(* IEC 61131-3 sources: s7-to-codesys/tests/POUs/Scenarios/FB_Sequencer_ScenarioTest, 7 files *)

(* ---- FB_Sequencer_ScenarioTest.decl.st ---- *)
// AUTO-GENERATED — не редактировать: s7conv gen-tests, сценарии scenarios/FB_Sequencer.csv
// Правка — в CSV (scenarios/README.md), затем python -m s7conv build-corpus.
// Назначение: тесты поведения сконвертированного FB_Sequencer по сценариям CSV (сценариев: 6, строк: 42):
//             один метод-тест на сценарий, строки — по порядку с моделируемым временем GVL_S7Clock.
//             Ожидаемые значения — из CSV (эталонные модели по описанию логики блока), не из
//             результата конвертации.
// Автор:      s7conv 0.1.0 (сгенерировано)
// Версия:     не указана
// Документ:   scenarios/README.md, docs/methodology.md, раздел «Проверка поведения»
FUNCTION_BLOCK FB_Sequencer_ScenarioTest EXTENDS coUnit.FB_TestSuite
VAR
    fbFullCycle : FB_Sequencer;  // свой экземпляр на сценарий
    xFullCycleDone : BOOL;  // сценарий выполнен (выполняется один раз)
    fbDrainTimeout : FB_Sequencer;  // свой экземпляр на сценарий
    xDrainTimeoutDone : BOOL;  // сценарий выполнен (выполняется один раз)
    fbAbortByStop : FB_Sequencer;  // свой экземпляр на сценарий
    xAbortByStopDone : BOOL;  // сценарий выполнен (выполняется один раз)
    fbPermissiveMissing : FB_Sequencer;  // свой экземпляр на сценарий
    xPermissiveMissingDone : BOOL;  // сценарий выполнен (выполняется один раз)
    fbDrainTimeoutBoundary : FB_Sequencer;  // свой экземпляр на сценарий
    xDrainTimeoutBoundaryDone : BOOL;  // сценарий выполнен (выполняется один раз)
    fbRefillTimeoutBoundary : FB_Sequencer;  // свой экземпляр на сценарий
    xRefillTimeoutBoundaryDone : BOOL;  // сценарий выполнен (выполняется один раз)
END_VAR

(* ---- AbortByStop.method.impl.st ---- *)
// AUTO-GENERATED — не редактировать: scenarios/FB_Sequencer.csv, сценарий AbortByStop
coUnit.TEST('AbortByStop');
IF NOT xAbortByStopDone THEN
    xAbortByStopDone := TRUE;
    GVL_S7Clock.xSimulation := TRUE;

    // #1, t = 0 мс — ожидание
    GVL_S7Clock.tSimNow := T#0MS;
    fbAbortByStop.start := FALSE;
    fbAbortByStop.stop := FALSE;
    fbAbortByStop.permissive := TRUE;
    fbAbortByStop.levelLow := FALSE;
    fbAbortByStop.levelHigh := FALSE;
    fbAbortByStop.reset := FALSE;
    fbAbortByStop.drainTimeout := T#60000MS;
    fbAbortByStop.airTime := T#30000MS;
    fbAbortByStop.washTime := T#40000MS;
    fbAbortByStop.refillTimeout := T#90000MS;
    fbAbortByStop();
    AssertEquals_INT(Expected := 0, Actual := fbAbortByStop.stepNo, Message := 'AbortByStop#1 stepNo');
    AssertEquals_BOOL(Expected := FALSE, Actual := fbAbortByStop.drainValve, Message := 'AbortByStop#1 drainValve');
    AssertEquals_BOOL(Expected := FALSE, Actual := fbAbortByStop.airBlower, Message := 'AbortByStop#1 airBlower');
    AssertEquals_BOOL(Expected := FALSE, Actual := fbAbortByStop.washPump, Message := 'AbortByStop#1 washPump');
    AssertEquals_BOOL(Expected := FALSE, Actual := fbAbortByStop.inletValve, Message := 'AbortByStop#1 inletValve');
    AssertEquals_BOOL(Expected := FALSE, Actual := fbAbortByStop.busy, Message := 'AbortByStop#1 busy');
    AssertEquals_BOOL(Expected := FALSE, Actual := fbAbortByStop.fault, Message := 'AbortByStop#1 fault');
    AssertEquals_INT(Expected := 0, Actual := fbAbortByStop.faultStep, Message := 'AbortByStop#1 faultStep');
    AssertEquals_DINT(Expected := 0, Actual := fbAbortByStop.cycleCount, Message := 'AbortByStop#1 cycleCount');
    AssertEquals_STRING(Expected := 'IDLE', Actual := fbAbortByStop.stepText, Message := 'AbortByStop#1 stepText');

    // #2, t = 1000 мс — пуск: опорожнение
    GVL_S7Clock.tSimNow := T#1000MS;
    fbAbortByStop.start := TRUE;
    fbAbortByStop();
    AssertEquals_INT(Expected := 10, Actual := fbAbortByStop.stepNo, Message := 'AbortByStop#2 stepNo');
    AssertEquals_BOOL(Expected := TRUE, Actual := fbAbortByStop.drainValve, Message := 'AbortByStop#2 drainValve');
    AssertEquals_BOOL(Expected := FALSE, Actual := fbAbortByStop.airBlower, Message := 'AbortByStop#2 airBlower');
    AssertEquals_BOOL(Expected := FALSE, Actual := fbAbortByStop.washPump, Message := 'AbortByStop#2 washPump');
    AssertEquals_BOOL(Expected := FALSE, Actual := fbAbortByStop.inletValve, Message := 'AbortByStop#2 inletValve');
    AssertEquals_BOOL(Expected := TRUE, Actual := fbAbortByStop.busy, Message := 'AbortByStop#2 busy');
    AssertEquals_BOOL(Expected := FALSE, Actual := fbAbortByStop.fault, Message := 'AbortByStop#2 fault');
    AssertEquals_INT(Expected := 0, Actual := fbAbortByStop.faultStep, Message := 'AbortByStop#2 faultStep');
    AssertEquals_DINT(Expected := 0, Actual := fbAbortByStop.cycleCount, Message := 'AbortByStop#2 cycleCount');
    AssertEquals_STRING(Expected := 'DRAIN', Actual := fbAbortByStop.stepText, Message := 'AbortByStop#2 stepText');

    // #3, t = 5000 мс — продувка с 5.0 с
    GVL_S7Clock.tSimNow := T#5000MS;
    fbAbortByStop.start := FALSE;
    fbAbortByStop.levelLow := TRUE;
    fbAbortByStop();
    AssertEquals_INT(Expected := 20, Actual := fbAbortByStop.stepNo, Message := 'AbortByStop#3 stepNo');
    AssertEquals_BOOL(Expected := FALSE, Actual := fbAbortByStop.drainValve, Message := 'AbortByStop#3 drainValve');
    AssertEquals_BOOL(Expected := TRUE, Actual := fbAbortByStop.airBlower, Message := 'AbortByStop#3 airBlower');
    AssertEquals_BOOL(Expected := FALSE, Actual := fbAbortByStop.washPump, Message := 'AbortByStop#3 washPump');
    AssertEquals_BOOL(Expected := FALSE, Actual := fbAbortByStop.inletValve, Message := 'AbortByStop#3 inletValve');
    AssertEquals_BOOL(Expected := TRUE, Actual := fbAbortByStop.busy, Message := 'AbortByStop#3 busy');
    AssertEquals_BOOL(Expected := FALSE, Actual := fbAbortByStop.fault, Message := 'AbortByStop#3 fault');
    AssertEquals_INT(Expected := 0, Actual := fbAbortByStop.faultStep, Message := 'AbortByStop#3 faultStep');
    AssertEquals_DINT(Expected := 0, Actual := fbAbortByStop.cycleCount, Message := 'AbortByStop#3 cycleCount');
    AssertEquals_STRING(Expected := 'AIR SCOUR', Actual := fbAbortByStop.stepText, Message := 'AbortByStop#3 stepText');

    // #4, t = 10000 мс — прерывание: ожидание, без аварии и без счёта
    GVL_S7Clock.tSimNow := T#10000MS;
    fbAbortByStop.stop := TRUE;
    fbAbortByStop();
    AssertEquals_INT(Expected := 0, Actual := fbAbortByStop.stepNo, Message := 'AbortByStop#4 stepNo');
    AssertEquals_BOOL(Expected := FALSE, Actual := fbAbortByStop.drainValve, Message := 'AbortByStop#4 drainValve');
    AssertEquals_BOOL(Expected := FALSE, Actual := fbAbortByStop.airBlower, Message := 'AbortByStop#4 airBlower');
    AssertEquals_BOOL(Expected := FALSE, Actual := fbAbortByStop.washPump, Message := 'AbortByStop#4 washPump');
    AssertEquals_BOOL(Expected := FALSE, Actual := fbAbortByStop.inletValve, Message := 'AbortByStop#4 inletValve');
    AssertEquals_BOOL(Expected := FALSE, Actual := fbAbortByStop.busy, Message := 'AbortByStop#4 busy');
    AssertEquals_BOOL(Expected := FALSE, Actual := fbAbortByStop.fault, Message := 'AbortByStop#4 fault');
    AssertEquals_INT(Expected := 0, Actual := fbAbortByStop.faultStep, Message := 'AbortByStop#4 faultStep');
    AssertEquals_DINT(Expected := 0, Actual := fbAbortByStop.cycleCount, Message := 'AbortByStop#4 cycleCount');
    AssertEquals_STRING(Expected := 'IDLE', Actual := fbAbortByStop.stepText, Message := 'AbortByStop#4 stepText');

    // #5, t = 11000 мс — фронт start при stop: не запускается
    GVL_S7Clock.tSimNow := T#11000MS;
    fbAbortByStop.start := TRUE;
    fbAbortByStop();
    AssertEquals_INT(Expected := 0, Actual := fbAbortByStop.stepNo, Message := 'AbortByStop#5 stepNo');
    AssertEquals_BOOL(Expected := FALSE, Actual := fbAbortByStop.drainValve, Message := 'AbortByStop#5 drainValve');
    AssertEquals_BOOL(Expected := FALSE, Actual := fbAbortByStop.airBlower, Message := 'AbortByStop#5 airBlower');
    AssertEquals_BOOL(Expected := FALSE, Actual := fbAbortByStop.washPump, Message := 'AbortByStop#5 washPump');
    AssertEquals_BOOL(Expected := FALSE, Actual := fbAbortByStop.inletValve, Message := 'AbortByStop#5 inletValve');
    AssertEquals_BOOL(Expected := FALSE, Actual := fbAbortByStop.busy, Message := 'AbortByStop#5 busy');
    AssertEquals_BOOL(Expected := FALSE, Actual := fbAbortByStop.fault, Message := 'AbortByStop#5 fault');
    AssertEquals_INT(Expected := 0, Actual := fbAbortByStop.faultStep, Message := 'AbortByStop#5 faultStep');
    AssertEquals_DINT(Expected := 0, Actual := fbAbortByStop.cycleCount, Message := 'AbortByStop#5 cycleCount');
    AssertEquals_STRING(Expected := 'IDLE', Actual := fbAbortByStop.stepText, Message := 'AbortByStop#5 stepText');

    // #6, t = 12000 мс — stop снят
    GVL_S7Clock.tSimNow := T#12000MS;
    fbAbortByStop.start := FALSE;
    fbAbortByStop.stop := FALSE;
    fbAbortByStop();
    AssertEquals_INT(Expected := 0, Actual := fbAbortByStop.stepNo, Message := 'AbortByStop#6 stepNo');
    AssertEquals_BOOL(Expected := FALSE, Actual := fbAbortByStop.drainValve, Message := 'AbortByStop#6 drainValve');
    AssertEquals_BOOL(Expected := FALSE, Actual := fbAbortByStop.airBlower, Message := 'AbortByStop#6 airBlower');
    AssertEquals_BOOL(Expected := FALSE, Actual := fbAbortByStop.washPump, Message := 'AbortByStop#6 washPump');
    AssertEquals_BOOL(Expected := FALSE, Actual := fbAbortByStop.inletValve, Message := 'AbortByStop#6 inletValve');
    AssertEquals_BOOL(Expected := FALSE, Actual := fbAbortByStop.busy, Message := 'AbortByStop#6 busy');
    AssertEquals_BOOL(Expected := FALSE, Actual := fbAbortByStop.fault, Message := 'AbortByStop#6 fault');
    AssertEquals_INT(Expected := 0, Actual := fbAbortByStop.faultStep, Message := 'AbortByStop#6 faultStep');
    AssertEquals_DINT(Expected := 0, Actual := fbAbortByStop.cycleCount, Message := 'AbortByStop#6 cycleCount');
    AssertEquals_STRING(Expected := 'IDLE', Actual := fbAbortByStop.stepText, Message := 'AbortByStop#6 stepText');

    // #7, t = 13000 мс — новый фронт start: опорожнение
    GVL_S7Clock.tSimNow := T#13000MS;
    fbAbortByStop.start := TRUE;
    fbAbortByStop();
    AssertEquals_INT(Expected := 10, Actual := fbAbortByStop.stepNo, Message := 'AbortByStop#7 stepNo');
    AssertEquals_BOOL(Expected := TRUE, Actual := fbAbortByStop.drainValve, Message := 'AbortByStop#7 drainValve');
    AssertEquals_BOOL(Expected := FALSE, Actual := fbAbortByStop.airBlower, Message := 'AbortByStop#7 airBlower');
    AssertEquals_BOOL(Expected := FALSE, Actual := fbAbortByStop.washPump, Message := 'AbortByStop#7 washPump');
    AssertEquals_BOOL(Expected := FALSE, Actual := fbAbortByStop.inletValve, Message := 'AbortByStop#7 inletValve');
    AssertEquals_BOOL(Expected := TRUE, Actual := fbAbortByStop.busy, Message := 'AbortByStop#7 busy');
    AssertEquals_BOOL(Expected := FALSE, Actual := fbAbortByStop.fault, Message := 'AbortByStop#7 fault');
    AssertEquals_INT(Expected := 0, Actual := fbAbortByStop.faultStep, Message := 'AbortByStop#7 faultStep');
    AssertEquals_DINT(Expected := 0, Actual := fbAbortByStop.cycleCount, Message := 'AbortByStop#7 cycleCount');
    AssertEquals_STRING(Expected := 'DRAIN', Actual := fbAbortByStop.stepText, Message := 'AbortByStop#7 stepText');

    GVL_S7Clock.xSimulation := FALSE;
END_IF
coUnit.TEST_FINISHED();

(* ---- DrainTimeout.method.impl.st ---- *)
// AUTO-GENERATED — не редактировать: scenarios/FB_Sequencer.csv, сценарий DrainTimeout
coUnit.TEST('DrainTimeout');
IF NOT xDrainTimeoutDone THEN
    xDrainTimeoutDone := TRUE;
    GVL_S7Clock.xSimulation := TRUE;

    // #1, t = 0 мс — ожидание
    GVL_S7Clock.tSimNow := T#0MS;
    fbDrainTimeout.start := FALSE;
    fbDrainTimeout.stop := FALSE;
    fbDrainTimeout.permissive := TRUE;
    fbDrainTimeout.levelLow := FALSE;
    fbDrainTimeout.levelHigh := FALSE;
    fbDrainTimeout.reset := FALSE;
    fbDrainTimeout.drainTimeout := T#60000MS;
    fbDrainTimeout.airTime := T#30000MS;
    fbDrainTimeout.washTime := T#40000MS;
    fbDrainTimeout.refillTimeout := T#90000MS;
    fbDrainTimeout();
    AssertEquals_INT(Expected := 0, Actual := fbDrainTimeout.stepNo, Message := 'DrainTimeout#1 stepNo');
    AssertEquals_BOOL(Expected := FALSE, Actual := fbDrainTimeout.drainValve, Message := 'DrainTimeout#1 drainValve');
    AssertEquals_BOOL(Expected := FALSE, Actual := fbDrainTimeout.airBlower, Message := 'DrainTimeout#1 airBlower');
    AssertEquals_BOOL(Expected := FALSE, Actual := fbDrainTimeout.washPump, Message := 'DrainTimeout#1 washPump');
    AssertEquals_BOOL(Expected := FALSE, Actual := fbDrainTimeout.inletValve, Message := 'DrainTimeout#1 inletValve');
    AssertEquals_BOOL(Expected := FALSE, Actual := fbDrainTimeout.busy, Message := 'DrainTimeout#1 busy');
    AssertEquals_BOOL(Expected := FALSE, Actual := fbDrainTimeout.fault, Message := 'DrainTimeout#1 fault');
    AssertEquals_INT(Expected := 0, Actual := fbDrainTimeout.faultStep, Message := 'DrainTimeout#1 faultStep');
    AssertEquals_DINT(Expected := 0, Actual := fbDrainTimeout.cycleCount, Message := 'DrainTimeout#1 cycleCount');
    AssertEquals_STRING(Expected := 'IDLE', Actual := fbDrainTimeout.stepText, Message := 'DrainTimeout#1 stepText');

    // #2, t = 1000 мс — пуск: опорожнение с 1.0 с
    GVL_S7Clock.tSimNow := T#1000MS;
    fbDrainTimeout.start := TRUE;
    fbDrainTimeout();
    AssertEquals_INT(Expected := 10, Actual := fbDrainTimeout.stepNo, Message := 'DrainTimeout#2 stepNo');
    AssertEquals_BOOL(Expected := TRUE, Actual := fbDrainTimeout.drainValve, Message := 'DrainTimeout#2 drainValve');
    AssertEquals_BOOL(Expected := FALSE, Actual := fbDrainTimeout.airBlower, Message := 'DrainTimeout#2 airBlower');
    AssertEquals_BOOL(Expected := FALSE, Actual := fbDrainTimeout.washPump, Message := 'DrainTimeout#2 washPump');
    AssertEquals_BOOL(Expected := FALSE, Actual := fbDrainTimeout.inletValve, Message := 'DrainTimeout#2 inletValve');
    AssertEquals_BOOL(Expected := TRUE, Actual := fbDrainTimeout.busy, Message := 'DrainTimeout#2 busy');
    AssertEquals_BOOL(Expected := FALSE, Actual := fbDrainTimeout.fault, Message := 'DrainTimeout#2 fault');
    AssertEquals_INT(Expected := 0, Actual := fbDrainTimeout.faultStep, Message := 'DrainTimeout#2 faultStep');
    AssertEquals_DINT(Expected := 0, Actual := fbDrainTimeout.cycleCount, Message := 'DrainTimeout#2 cycleCount');
    AssertEquals_STRING(Expected := 'DRAIN', Actual := fbDrainTimeout.stepText, Message := 'DrainTimeout#2 stepText');

    // #3, t = 60800 мс — 59.8 с < 60 с: опорожнение
    GVL_S7Clock.tSimNow := T#60800MS;
    fbDrainTimeout.start := FALSE;
    fbDrainTimeout();
    AssertEquals_INT(Expected := 10, Actual := fbDrainTimeout.stepNo, Message := 'DrainTimeout#3 stepNo');
    AssertEquals_BOOL(Expected := TRUE, Actual := fbDrainTimeout.drainValve, Message := 'DrainTimeout#3 drainValve');
    AssertEquals_BOOL(Expected := FALSE, Actual := fbDrainTimeout.airBlower, Message := 'DrainTimeout#3 airBlower');
    AssertEquals_BOOL(Expected := FALSE, Actual := fbDrainTimeout.washPump, Message := 'DrainTimeout#3 washPump');
    AssertEquals_BOOL(Expected := FALSE, Actual := fbDrainTimeout.inletValve, Message := 'DrainTimeout#3 inletValve');
    AssertEquals_BOOL(Expected := TRUE, Actual := fbDrainTimeout.busy, Message := 'DrainTimeout#3 busy');
    AssertEquals_BOOL(Expected := FALSE, Actual := fbDrainTimeout.fault, Message := 'DrainTimeout#3 fault');
    AssertEquals_INT(Expected := 0, Actual := fbDrainTimeout.faultStep, Message := 'DrainTimeout#3 faultStep');
    AssertEquals_DINT(Expected := 0, Actual := fbDrainTimeout.cycleCount, Message := 'DrainTimeout#3 cycleCount');
    AssertEquals_STRING(Expected := 'DRAIN', Actual := fbDrainTimeout.stepText, Message := 'DrainTimeout#3 stepText');

    // #4, t = 61200 мс — 60.2 с: авария на шаге 10, всё закрыто
    GVL_S7Clock.tSimNow := T#61200MS;
    fbDrainTimeout();
    AssertEquals_INT(Expected := 90, Actual := fbDrainTimeout.stepNo, Message := 'DrainTimeout#4 stepNo');
    AssertEquals_BOOL(Expected := FALSE, Actual := fbDrainTimeout.drainValve, Message := 'DrainTimeout#4 drainValve');
    AssertEquals_BOOL(Expected := FALSE, Actual := fbDrainTimeout.airBlower, Message := 'DrainTimeout#4 airBlower');
    AssertEquals_BOOL(Expected := FALSE, Actual := fbDrainTimeout.washPump, Message := 'DrainTimeout#4 washPump');
    AssertEquals_BOOL(Expected := FALSE, Actual := fbDrainTimeout.inletValve, Message := 'DrainTimeout#4 inletValve');
    AssertEquals_BOOL(Expected := FALSE, Actual := fbDrainTimeout.busy, Message := 'DrainTimeout#4 busy');
    AssertEquals_BOOL(Expected := TRUE, Actual := fbDrainTimeout.fault, Message := 'DrainTimeout#4 fault');
    AssertEquals_INT(Expected := 10, Actual := fbDrainTimeout.faultStep, Message := 'DrainTimeout#4 faultStep');
    AssertEquals_DINT(Expected := 0, Actual := fbDrainTimeout.cycleCount, Message := 'DrainTimeout#4 cycleCount');
    AssertEquals_STRING(Expected := 'FAULT', Actual := fbDrainTimeout.stepText, Message := 'DrainTimeout#4 stepText');

    // #5, t = 65000 мс — пуск во время аварии не действует
    GVL_S7Clock.tSimNow := T#65000MS;
    fbDrainTimeout.start := TRUE;
    fbDrainTimeout();
    AssertEquals_INT(Expected := 90, Actual := fbDrainTimeout.stepNo, Message := 'DrainTimeout#5 stepNo');
    AssertEquals_BOOL(Expected := FALSE, Actual := fbDrainTimeout.drainValve, Message := 'DrainTimeout#5 drainValve');
    AssertEquals_BOOL(Expected := FALSE, Actual := fbDrainTimeout.airBlower, Message := 'DrainTimeout#5 airBlower');
    AssertEquals_BOOL(Expected := FALSE, Actual := fbDrainTimeout.washPump, Message := 'DrainTimeout#5 washPump');
    AssertEquals_BOOL(Expected := FALSE, Actual := fbDrainTimeout.inletValve, Message := 'DrainTimeout#5 inletValve');
    AssertEquals_BOOL(Expected := FALSE, Actual := fbDrainTimeout.busy, Message := 'DrainTimeout#5 busy');
    AssertEquals_BOOL(Expected := TRUE, Actual := fbDrainTimeout.fault, Message := 'DrainTimeout#5 fault');
    AssertEquals_INT(Expected := 10, Actual := fbDrainTimeout.faultStep, Message := 'DrainTimeout#5 faultStep');
    AssertEquals_DINT(Expected := 0, Actual := fbDrainTimeout.cycleCount, Message := 'DrainTimeout#5 cycleCount');
    AssertEquals_STRING(Expected := 'FAULT', Actual := fbDrainTimeout.stepText, Message := 'DrainTimeout#5 stepText');

    // #6, t = 70000 мс — сброс: ожидание, faultStep 0
    GVL_S7Clock.tSimNow := T#70000MS;
    fbDrainTimeout.start := FALSE;
    fbDrainTimeout.reset := TRUE;
    fbDrainTimeout();
    AssertEquals_INT(Expected := 0, Actual := fbDrainTimeout.stepNo, Message := 'DrainTimeout#6 stepNo');
    AssertEquals_BOOL(Expected := FALSE, Actual := fbDrainTimeout.drainValve, Message := 'DrainTimeout#6 drainValve');
    AssertEquals_BOOL(Expected := FALSE, Actual := fbDrainTimeout.airBlower, Message := 'DrainTimeout#6 airBlower');
    AssertEquals_BOOL(Expected := FALSE, Actual := fbDrainTimeout.washPump, Message := 'DrainTimeout#6 washPump');
    AssertEquals_BOOL(Expected := FALSE, Actual := fbDrainTimeout.inletValve, Message := 'DrainTimeout#6 inletValve');
    AssertEquals_BOOL(Expected := FALSE, Actual := fbDrainTimeout.busy, Message := 'DrainTimeout#6 busy');
    AssertEquals_BOOL(Expected := FALSE, Actual := fbDrainTimeout.fault, Message := 'DrainTimeout#6 fault');
    AssertEquals_INT(Expected := 0, Actual := fbDrainTimeout.faultStep, Message := 'DrainTimeout#6 faultStep');
    AssertEquals_DINT(Expected := 0, Actual := fbDrainTimeout.cycleCount, Message := 'DrainTimeout#6 cycleCount');
    AssertEquals_STRING(Expected := 'IDLE', Actual := fbDrainTimeout.stepText, Message := 'DrainTimeout#6 stepText');

    // #7, t = 71000 мс — ожидание
    GVL_S7Clock.tSimNow := T#71000MS;
    fbDrainTimeout.reset := FALSE;
    fbDrainTimeout();
    AssertEquals_INT(Expected := 0, Actual := fbDrainTimeout.stepNo, Message := 'DrainTimeout#7 stepNo');
    AssertEquals_BOOL(Expected := FALSE, Actual := fbDrainTimeout.drainValve, Message := 'DrainTimeout#7 drainValve');
    AssertEquals_BOOL(Expected := FALSE, Actual := fbDrainTimeout.airBlower, Message := 'DrainTimeout#7 airBlower');
    AssertEquals_BOOL(Expected := FALSE, Actual := fbDrainTimeout.washPump, Message := 'DrainTimeout#7 washPump');
    AssertEquals_BOOL(Expected := FALSE, Actual := fbDrainTimeout.inletValve, Message := 'DrainTimeout#7 inletValve');
    AssertEquals_BOOL(Expected := FALSE, Actual := fbDrainTimeout.busy, Message := 'DrainTimeout#7 busy');
    AssertEquals_BOOL(Expected := FALSE, Actual := fbDrainTimeout.fault, Message := 'DrainTimeout#7 fault');
    AssertEquals_INT(Expected := 0, Actual := fbDrainTimeout.faultStep, Message := 'DrainTimeout#7 faultStep');
    AssertEquals_DINT(Expected := 0, Actual := fbDrainTimeout.cycleCount, Message := 'DrainTimeout#7 cycleCount');
    AssertEquals_STRING(Expected := 'IDLE', Actual := fbDrainTimeout.stepText, Message := 'DrainTimeout#7 stepText');

    GVL_S7Clock.xSimulation := FALSE;
END_IF
coUnit.TEST_FINISHED();

(* ---- DrainTimeoutBoundary.method.impl.st ---- *)
// AUTO-GENERATED — не редактировать: scenarios/FB_Sequencer.csv, сценарий DrainTimeoutBoundary
coUnit.TEST('DrainTimeoutBoundary');
IF NOT xDrainTimeoutBoundaryDone THEN
    xDrainTimeoutBoundaryDone := TRUE;
    GVL_S7Clock.xSimulation := TRUE;

    // #1, t = 0 мс — пуск в первом вызове: опорожнение с 0 с
    GVL_S7Clock.tSimNow := T#0MS;
    fbDrainTimeoutBoundary.start := TRUE;
    fbDrainTimeoutBoundary.stop := FALSE;
    fbDrainTimeoutBoundary.permissive := TRUE;
    fbDrainTimeoutBoundary.levelLow := FALSE;
    fbDrainTimeoutBoundary.levelHigh := FALSE;
    fbDrainTimeoutBoundary.reset := FALSE;
    fbDrainTimeoutBoundary.drainTimeout := T#60000MS;
    fbDrainTimeoutBoundary.airTime := T#30000MS;
    fbDrainTimeoutBoundary.washTime := T#40000MS;
    fbDrainTimeoutBoundary.refillTimeout := T#90000MS;
    fbDrainTimeoutBoundary();
    AssertEquals_INT(Expected := 10,
                     Actual := fbDrainTimeoutBoundary.stepNo,
                     Message := 'DrainTimeoutBoundary#1 stepNo');
    AssertEquals_BOOL(Expected := TRUE,
                      Actual := fbDrainTimeoutBoundary.drainValve,
                      Message := 'DrainTimeoutBoundary#1 drainValve');
    AssertEquals_BOOL(Expected := FALSE,
                      Actual := fbDrainTimeoutBoundary.airBlower,
                      Message := 'DrainTimeoutBoundary#1 airBlower');
    AssertEquals_BOOL(Expected := FALSE,
                      Actual := fbDrainTimeoutBoundary.washPump,
                      Message := 'DrainTimeoutBoundary#1 washPump');
    AssertEquals_BOOL(Expected := FALSE,
                      Actual := fbDrainTimeoutBoundary.inletValve,
                      Message := 'DrainTimeoutBoundary#1 inletValve');
    AssertEquals_BOOL(Expected := TRUE,
                      Actual := fbDrainTimeoutBoundary.busy,
                      Message := 'DrainTimeoutBoundary#1 busy');
    AssertEquals_BOOL(Expected := FALSE,
                      Actual := fbDrainTimeoutBoundary.fault,
                      Message := 'DrainTimeoutBoundary#1 fault');
    AssertEquals_INT(Expected := 0,
                     Actual := fbDrainTimeoutBoundary.faultStep,
                     Message := 'DrainTimeoutBoundary#1 faultStep');
    AssertEquals_DINT(Expected := 0,
                      Actual := fbDrainTimeoutBoundary.cycleCount,
                      Message := 'DrainTimeoutBoundary#1 cycleCount');
    AssertEquals_STRING(Expected := 'DRAIN',
                        Actual := fbDrainTimeoutBoundary.stepText,
                        Message := 'DrainTimeoutBoundary#1 stepText');

    // #2, t = 59800 мс — 59.8 с: опорожнение
    GVL_S7Clock.tSimNow := T#59800MS;
    fbDrainTimeoutBoundary.start := FALSE;
    fbDrainTimeoutBoundary();
    AssertEquals_INT(Expected := 10,
                     Actual := fbDrainTimeoutBoundary.stepNo,
                     Message := 'DrainTimeoutBoundary#2 stepNo');
    AssertEquals_BOOL(Expected := TRUE,
                      Actual := fbDrainTimeoutBoundary.drainValve,
                      Message := 'DrainTimeoutBoundary#2 drainValve');
    AssertEquals_BOOL(Expected := FALSE,
                      Actual := fbDrainTimeoutBoundary.airBlower,
                      Message := 'DrainTimeoutBoundary#2 airBlower');
    AssertEquals_BOOL(Expected := FALSE,
                      Actual := fbDrainTimeoutBoundary.washPump,
                      Message := 'DrainTimeoutBoundary#2 washPump');
    AssertEquals_BOOL(Expected := FALSE,
                      Actual := fbDrainTimeoutBoundary.inletValve,
                      Message := 'DrainTimeoutBoundary#2 inletValve');
    AssertEquals_BOOL(Expected := TRUE,
                      Actual := fbDrainTimeoutBoundary.busy,
                      Message := 'DrainTimeoutBoundary#2 busy');
    AssertEquals_BOOL(Expected := FALSE,
                      Actual := fbDrainTimeoutBoundary.fault,
                      Message := 'DrainTimeoutBoundary#2 fault');
    AssertEquals_INT(Expected := 0,
                     Actual := fbDrainTimeoutBoundary.faultStep,
                     Message := 'DrainTimeoutBoundary#2 faultStep');
    AssertEquals_DINT(Expected := 0,
                      Actual := fbDrainTimeoutBoundary.cycleCount,
                      Message := 'DrainTimeoutBoundary#2 cycleCount');
    AssertEquals_STRING(Expected := 'DRAIN',
                        Actual := fbDrainTimeoutBoundary.stepText,
                        Message := 'DrainTimeoutBoundary#2 stepText');

    // #3, t = 60000 мс, на пороге таймера — 60.0 с = drainTimeout: авария
    GVL_S7Clock.tSimNow := T#60000MS;
    fbDrainTimeoutBoundary();
    AssertEquals_INT(Expected := 90,
                     Actual := fbDrainTimeoutBoundary.stepNo,
                     Message := 'DrainTimeoutBoundary#3 stepNo');
    AssertEquals_BOOL(Expected := FALSE,
                      Actual := fbDrainTimeoutBoundary.drainValve,
                      Message := 'DrainTimeoutBoundary#3 drainValve');
    AssertEquals_BOOL(Expected := FALSE,
                      Actual := fbDrainTimeoutBoundary.airBlower,
                      Message := 'DrainTimeoutBoundary#3 airBlower');
    AssertEquals_BOOL(Expected := FALSE,
                      Actual := fbDrainTimeoutBoundary.washPump,
                      Message := 'DrainTimeoutBoundary#3 washPump');
    AssertEquals_BOOL(Expected := FALSE,
                      Actual := fbDrainTimeoutBoundary.inletValve,
                      Message := 'DrainTimeoutBoundary#3 inletValve');
    AssertEquals_BOOL(Expected := FALSE,
                      Actual := fbDrainTimeoutBoundary.busy,
                      Message := 'DrainTimeoutBoundary#3 busy');
    AssertEquals_BOOL(Expected := TRUE,
                      Actual := fbDrainTimeoutBoundary.fault,
                      Message := 'DrainTimeoutBoundary#3 fault');
    AssertEquals_INT(Expected := 10,
                     Actual := fbDrainTimeoutBoundary.faultStep,
                     Message := 'DrainTimeoutBoundary#3 faultStep');
    AssertEquals_DINT(Expected := 0,
                      Actual := fbDrainTimeoutBoundary.cycleCount,
                      Message := 'DrainTimeoutBoundary#3 cycleCount');
    AssertEquals_STRING(Expected := 'FAULT',
                        Actual := fbDrainTimeoutBoundary.stepText,
                        Message := 'DrainTimeoutBoundary#3 stepText');

    // #4, t = 60200 мс — авария
    GVL_S7Clock.tSimNow := T#60200MS;
    fbDrainTimeoutBoundary();
    AssertEquals_INT(Expected := 90,
                     Actual := fbDrainTimeoutBoundary.stepNo,
                     Message := 'DrainTimeoutBoundary#4 stepNo');
    AssertEquals_BOOL(Expected := FALSE,
                      Actual := fbDrainTimeoutBoundary.drainValve,
                      Message := 'DrainTimeoutBoundary#4 drainValve');
    AssertEquals_BOOL(Expected := FALSE,
                      Actual := fbDrainTimeoutBoundary.airBlower,
                      Message := 'DrainTimeoutBoundary#4 airBlower');
    AssertEquals_BOOL(Expected := FALSE,
                      Actual := fbDrainTimeoutBoundary.washPump,
                      Message := 'DrainTimeoutBoundary#4 washPump');
    AssertEquals_BOOL(Expected := FALSE,
                      Actual := fbDrainTimeoutBoundary.inletValve,
                      Message := 'DrainTimeoutBoundary#4 inletValve');
    AssertEquals_BOOL(Expected := FALSE,
                      Actual := fbDrainTimeoutBoundary.busy,
                      Message := 'DrainTimeoutBoundary#4 busy');
    AssertEquals_BOOL(Expected := TRUE,
                      Actual := fbDrainTimeoutBoundary.fault,
                      Message := 'DrainTimeoutBoundary#4 fault');
    AssertEquals_INT(Expected := 10,
                     Actual := fbDrainTimeoutBoundary.faultStep,
                     Message := 'DrainTimeoutBoundary#4 faultStep');
    AssertEquals_DINT(Expected := 0,
                      Actual := fbDrainTimeoutBoundary.cycleCount,
                      Message := 'DrainTimeoutBoundary#4 cycleCount');
    AssertEquals_STRING(Expected := 'FAULT',
                        Actual := fbDrainTimeoutBoundary.stepText,
                        Message := 'DrainTimeoutBoundary#4 stepText');

    GVL_S7Clock.xSimulation := FALSE;
END_IF
coUnit.TEST_FINISHED();

(* ---- FullCycle.method.impl.st ---- *)
// AUTO-GENERATED — не редактировать: scenarios/FB_Sequencer.csv, сценарий FullCycle
coUnit.TEST('FullCycle');
IF NOT xFullCycleDone THEN
    xFullCycleDone := TRUE;
    GVL_S7Clock.xSimulation := TRUE;

    // #1, t = 0 мс — ожидание
    GVL_S7Clock.tSimNow := T#0MS;
    fbFullCycle.start := FALSE;
    fbFullCycle.stop := FALSE;
    fbFullCycle.permissive := TRUE;
    fbFullCycle.levelLow := FALSE;
    fbFullCycle.levelHigh := FALSE;
    fbFullCycle.reset := FALSE;
    fbFullCycle.drainTimeout := T#60000MS;
    fbFullCycle.airTime := T#30000MS;
    fbFullCycle.washTime := T#40000MS;
    fbFullCycle.refillTimeout := T#90000MS;
    fbFullCycle();
    AssertEquals_INT(Expected := 0, Actual := fbFullCycle.stepNo, Message := 'FullCycle#1 stepNo');
    AssertEquals_BOOL(Expected := FALSE, Actual := fbFullCycle.drainValve, Message := 'FullCycle#1 drainValve');
    AssertEquals_BOOL(Expected := FALSE, Actual := fbFullCycle.airBlower, Message := 'FullCycle#1 airBlower');
    AssertEquals_BOOL(Expected := FALSE, Actual := fbFullCycle.washPump, Message := 'FullCycle#1 washPump');
    AssertEquals_BOOL(Expected := FALSE, Actual := fbFullCycle.inletValve, Message := 'FullCycle#1 inletValve');
    AssertEquals_BOOL(Expected := FALSE, Actual := fbFullCycle.busy, Message := 'FullCycle#1 busy');
    AssertEquals_BOOL(Expected := FALSE, Actual := fbFullCycle.fault, Message := 'FullCycle#1 fault');
    AssertEquals_INT(Expected := 0, Actual := fbFullCycle.faultStep, Message := 'FullCycle#1 faultStep');
    AssertEquals_DINT(Expected := 0, Actual := fbFullCycle.cycleCount, Message := 'FullCycle#1 cycleCount');
    AssertEquals_STRING(Expected := 'IDLE', Actual := fbFullCycle.stepText, Message := 'FullCycle#1 stepText');

    // #2, t = 1000 мс — пуск: опорожнение, шаг 10 с 1.0 с
    GVL_S7Clock.tSimNow := T#1000MS;
    fbFullCycle.start := TRUE;
    fbFullCycle();
    AssertEquals_INT(Expected := 10, Actual := fbFullCycle.stepNo, Message := 'FullCycle#2 stepNo');
    AssertEquals_BOOL(Expected := TRUE, Actual := fbFullCycle.drainValve, Message := 'FullCycle#2 drainValve');
    AssertEquals_BOOL(Expected := FALSE, Actual := fbFullCycle.airBlower, Message := 'FullCycle#2 airBlower');
    AssertEquals_BOOL(Expected := FALSE, Actual := fbFullCycle.washPump, Message := 'FullCycle#2 washPump');
    AssertEquals_BOOL(Expected := FALSE, Actual := fbFullCycle.inletValve, Message := 'FullCycle#2 inletValve');
    AssertEquals_BOOL(Expected := TRUE, Actual := fbFullCycle.busy, Message := 'FullCycle#2 busy');
    AssertEquals_BOOL(Expected := FALSE, Actual := fbFullCycle.fault, Message := 'FullCycle#2 fault');
    AssertEquals_INT(Expected := 0, Actual := fbFullCycle.faultStep, Message := 'FullCycle#2 faultStep');
    AssertEquals_DINT(Expected := 0, Actual := fbFullCycle.cycleCount, Message := 'FullCycle#2 cycleCount');
    AssertEquals_STRING(Expected := 'DRAIN', Actual := fbFullCycle.stepText, Message := 'FullCycle#2 stepText');

    // #3, t = 1500 мс — опорожнение
    GVL_S7Clock.tSimNow := T#1500MS;
    fbFullCycle.start := FALSE;
    fbFullCycle();
    AssertEquals_INT(Expected := 10, Actual := fbFullCycle.stepNo, Message := 'FullCycle#3 stepNo');
    AssertEquals_BOOL(Expected := TRUE, Actual := fbFullCycle.drainValve, Message := 'FullCycle#3 drainValve');
    AssertEquals_BOOL(Expected := FALSE, Actual := fbFullCycle.airBlower, Message := 'FullCycle#3 airBlower');
    AssertEquals_BOOL(Expected := FALSE, Actual := fbFullCycle.washPump, Message := 'FullCycle#3 washPump');
    AssertEquals_BOOL(Expected := FALSE, Actual := fbFullCycle.inletValve, Message := 'FullCycle#3 inletValve');
    AssertEquals_BOOL(Expected := TRUE, Actual := fbFullCycle.busy, Message := 'FullCycle#3 busy');
    AssertEquals_BOOL(Expected := FALSE, Actual := fbFullCycle.fault, Message := 'FullCycle#3 fault');
    AssertEquals_INT(Expected := 0, Actual := fbFullCycle.faultStep, Message := 'FullCycle#3 faultStep');
    AssertEquals_DINT(Expected := 0, Actual := fbFullCycle.cycleCount, Message := 'FullCycle#3 cycleCount');
    AssertEquals_STRING(Expected := 'DRAIN', Actual := fbFullCycle.stepText, Message := 'FullCycle#3 stepText');

    // #4, t = 21000 мс — фильтр опорожнён: продувка, шаг 20 с 21.0 с
    GVL_S7Clock.tSimNow := T#21000MS;
    fbFullCycle.levelLow := TRUE;
    fbFullCycle();
    AssertEquals_INT(Expected := 20, Actual := fbFullCycle.stepNo, Message := 'FullCycle#4 stepNo');
    AssertEquals_BOOL(Expected := FALSE, Actual := fbFullCycle.drainValve, Message := 'FullCycle#4 drainValve');
    AssertEquals_BOOL(Expected := TRUE, Actual := fbFullCycle.airBlower, Message := 'FullCycle#4 airBlower');
    AssertEquals_BOOL(Expected := FALSE, Actual := fbFullCycle.washPump, Message := 'FullCycle#4 washPump');
    AssertEquals_BOOL(Expected := FALSE, Actual := fbFullCycle.inletValve, Message := 'FullCycle#4 inletValve');
    AssertEquals_BOOL(Expected := TRUE, Actual := fbFullCycle.busy, Message := 'FullCycle#4 busy');
    AssertEquals_BOOL(Expected := FALSE, Actual := fbFullCycle.fault, Message := 'FullCycle#4 fault');
    AssertEquals_INT(Expected := 0, Actual := fbFullCycle.faultStep, Message := 'FullCycle#4 faultStep');
    AssertEquals_DINT(Expected := 0, Actual := fbFullCycle.cycleCount, Message := 'FullCycle#4 cycleCount');
    AssertEquals_STRING(Expected := 'AIR SCOUR', Actual := fbFullCycle.stepText, Message := 'FullCycle#4 stepText');

    // #5, t = 50800 мс — продувка 29.8 с < 30 с
    GVL_S7Clock.tSimNow := T#50800MS;
    fbFullCycle();
    AssertEquals_INT(Expected := 20, Actual := fbFullCycle.stepNo, Message := 'FullCycle#5 stepNo');
    AssertEquals_BOOL(Expected := FALSE, Actual := fbFullCycle.drainValve, Message := 'FullCycle#5 drainValve');
    AssertEquals_BOOL(Expected := TRUE, Actual := fbFullCycle.airBlower, Message := 'FullCycle#5 airBlower');
    AssertEquals_BOOL(Expected := FALSE, Actual := fbFullCycle.washPump, Message := 'FullCycle#5 washPump');
    AssertEquals_BOOL(Expected := FALSE, Actual := fbFullCycle.inletValve, Message := 'FullCycle#5 inletValve');
    AssertEquals_BOOL(Expected := TRUE, Actual := fbFullCycle.busy, Message := 'FullCycle#5 busy');
    AssertEquals_BOOL(Expected := FALSE, Actual := fbFullCycle.fault, Message := 'FullCycle#5 fault');
    AssertEquals_INT(Expected := 0, Actual := fbFullCycle.faultStep, Message := 'FullCycle#5 faultStep');
    AssertEquals_DINT(Expected := 0, Actual := fbFullCycle.cycleCount, Message := 'FullCycle#5 cycleCount');
    AssertEquals_STRING(Expected := 'AIR SCOUR', Actual := fbFullCycle.stepText, Message := 'FullCycle#5 stepText');

    // #6, t = 51200 мс — 30.2 с: промывка, шаг 30 с 51.2 с
    GVL_S7Clock.tSimNow := T#51200MS;
    fbFullCycle();
    AssertEquals_INT(Expected := 30, Actual := fbFullCycle.stepNo, Message := 'FullCycle#6 stepNo');
    AssertEquals_BOOL(Expected := TRUE, Actual := fbFullCycle.drainValve, Message := 'FullCycle#6 drainValve');
    AssertEquals_BOOL(Expected := FALSE, Actual := fbFullCycle.airBlower, Message := 'FullCycle#6 airBlower');
    AssertEquals_BOOL(Expected := TRUE, Actual := fbFullCycle.washPump, Message := 'FullCycle#6 washPump');
    AssertEquals_BOOL(Expected := FALSE, Actual := fbFullCycle.inletValve, Message := 'FullCycle#6 inletValve');
    AssertEquals_BOOL(Expected := TRUE, Actual := fbFullCycle.busy, Message := 'FullCycle#6 busy');
    AssertEquals_BOOL(Expected := FALSE, Actual := fbFullCycle.fault, Message := 'FullCycle#6 fault');
    AssertEquals_INT(Expected := 0, Actual := fbFullCycle.faultStep, Message := 'FullCycle#6 faultStep');
    AssertEquals_DINT(Expected := 0, Actual := fbFullCycle.cycleCount, Message := 'FullCycle#6 cycleCount');
    AssertEquals_STRING(Expected := 'BACKWASH', Actual := fbFullCycle.stepText, Message := 'FullCycle#6 stepText');

    // #7, t = 91000 мс — промывка 39.8 с < 40 с
    GVL_S7Clock.tSimNow := T#91000MS;
    fbFullCycle.levelLow := FALSE;
    fbFullCycle();
    AssertEquals_INT(Expected := 30, Actual := fbFullCycle.stepNo, Message := 'FullCycle#7 stepNo');
    AssertEquals_BOOL(Expected := TRUE, Actual := fbFullCycle.drainValve, Message := 'FullCycle#7 drainValve');
    AssertEquals_BOOL(Expected := FALSE, Actual := fbFullCycle.airBlower, Message := 'FullCycle#7 airBlower');
    AssertEquals_BOOL(Expected := TRUE, Actual := fbFullCycle.washPump, Message := 'FullCycle#7 washPump');
    AssertEquals_BOOL(Expected := FALSE, Actual := fbFullCycle.inletValve, Message := 'FullCycle#7 inletValve');
    AssertEquals_BOOL(Expected := TRUE, Actual := fbFullCycle.busy, Message := 'FullCycle#7 busy');
    AssertEquals_BOOL(Expected := FALSE, Actual := fbFullCycle.fault, Message := 'FullCycle#7 fault');
    AssertEquals_INT(Expected := 0, Actual := fbFullCycle.faultStep, Message := 'FullCycle#7 faultStep');
    AssertEquals_DINT(Expected := 0, Actual := fbFullCycle.cycleCount, Message := 'FullCycle#7 cycleCount');
    AssertEquals_STRING(Expected := 'BACKWASH', Actual := fbFullCycle.stepText, Message := 'FullCycle#7 stepText');

    // #8, t = 91400 мс — 40.2 с: заполнение, шаг 40 с 91.4 с
    GVL_S7Clock.tSimNow := T#91400MS;
    fbFullCycle();
    AssertEquals_INT(Expected := 40, Actual := fbFullCycle.stepNo, Message := 'FullCycle#8 stepNo');
    AssertEquals_BOOL(Expected := FALSE, Actual := fbFullCycle.drainValve, Message := 'FullCycle#8 drainValve');
    AssertEquals_BOOL(Expected := FALSE, Actual := fbFullCycle.airBlower, Message := 'FullCycle#8 airBlower');
    AssertEquals_BOOL(Expected := FALSE, Actual := fbFullCycle.washPump, Message := 'FullCycle#8 washPump');
    AssertEquals_BOOL(Expected := TRUE, Actual := fbFullCycle.inletValve, Message := 'FullCycle#8 inletValve');
    AssertEquals_BOOL(Expected := TRUE, Actual := fbFullCycle.busy, Message := 'FullCycle#8 busy');
    AssertEquals_BOOL(Expected := FALSE, Actual := fbFullCycle.fault, Message := 'FullCycle#8 fault');
    AssertEquals_INT(Expected := 0, Actual := fbFullCycle.faultStep, Message := 'FullCycle#8 faultStep');
    AssertEquals_DINT(Expected := 0, Actual := fbFullCycle.cycleCount, Message := 'FullCycle#8 cycleCount');
    AssertEquals_STRING(Expected := 'REFILL', Actual := fbFullCycle.stepText, Message := 'FullCycle#8 stepText');

    // #9, t = 150000 мс — заполнение 58.6 с, уровня нет
    GVL_S7Clock.tSimNow := T#150000MS;
    fbFullCycle();
    AssertEquals_INT(Expected := 40, Actual := fbFullCycle.stepNo, Message := 'FullCycle#9 stepNo');
    AssertEquals_BOOL(Expected := FALSE, Actual := fbFullCycle.drainValve, Message := 'FullCycle#9 drainValve');
    AssertEquals_BOOL(Expected := FALSE, Actual := fbFullCycle.airBlower, Message := 'FullCycle#9 airBlower');
    AssertEquals_BOOL(Expected := FALSE, Actual := fbFullCycle.washPump, Message := 'FullCycle#9 washPump');
    AssertEquals_BOOL(Expected := TRUE, Actual := fbFullCycle.inletValve, Message := 'FullCycle#9 inletValve');
    AssertEquals_BOOL(Expected := TRUE, Actual := fbFullCycle.busy, Message := 'FullCycle#9 busy');
    AssertEquals_BOOL(Expected := FALSE, Actual := fbFullCycle.fault, Message := 'FullCycle#9 fault');
    AssertEquals_INT(Expected := 0, Actual := fbFullCycle.faultStep, Message := 'FullCycle#9 faultStep');
    AssertEquals_DINT(Expected := 0, Actual := fbFullCycle.cycleCount, Message := 'FullCycle#9 cycleCount');
    AssertEquals_STRING(Expected := 'REFILL', Actual := fbFullCycle.stepText, Message := 'FullCycle#9 stepText');

    // #10, t = 160000 мс — фильтр заполнен: цикл №1 завершён
    GVL_S7Clock.tSimNow := T#160000MS;
    fbFullCycle.levelHigh := TRUE;
    fbFullCycle();
    AssertEquals_INT(Expected := 0, Actual := fbFullCycle.stepNo, Message := 'FullCycle#10 stepNo');
    AssertEquals_BOOL(Expected := FALSE, Actual := fbFullCycle.drainValve, Message := 'FullCycle#10 drainValve');
    AssertEquals_BOOL(Expected := FALSE, Actual := fbFullCycle.airBlower, Message := 'FullCycle#10 airBlower');
    AssertEquals_BOOL(Expected := FALSE, Actual := fbFullCycle.washPump, Message := 'FullCycle#10 washPump');
    AssertEquals_BOOL(Expected := FALSE, Actual := fbFullCycle.inletValve, Message := 'FullCycle#10 inletValve');
    AssertEquals_BOOL(Expected := FALSE, Actual := fbFullCycle.busy, Message := 'FullCycle#10 busy');
    AssertEquals_BOOL(Expected := FALSE, Actual := fbFullCycle.fault, Message := 'FullCycle#10 fault');
    AssertEquals_INT(Expected := 0, Actual := fbFullCycle.faultStep, Message := 'FullCycle#10 faultStep');
    AssertEquals_DINT(Expected := 1, Actual := fbFullCycle.cycleCount, Message := 'FullCycle#10 cycleCount');
    AssertEquals_STRING(Expected := 'IDLE', Actual := fbFullCycle.stepText, Message := 'FullCycle#10 stepText');

    // #11, t = 161000 мс — ожидание, повторного пуска без фронта start нет
    GVL_S7Clock.tSimNow := T#161000MS;
    fbFullCycle();
    AssertEquals_INT(Expected := 0, Actual := fbFullCycle.stepNo, Message := 'FullCycle#11 stepNo');
    AssertEquals_BOOL(Expected := FALSE, Actual := fbFullCycle.drainValve, Message := 'FullCycle#11 drainValve');
    AssertEquals_BOOL(Expected := FALSE, Actual := fbFullCycle.airBlower, Message := 'FullCycle#11 airBlower');
    AssertEquals_BOOL(Expected := FALSE, Actual := fbFullCycle.washPump, Message := 'FullCycle#11 washPump');
    AssertEquals_BOOL(Expected := FALSE, Actual := fbFullCycle.inletValve, Message := 'FullCycle#11 inletValve');
    AssertEquals_BOOL(Expected := FALSE, Actual := fbFullCycle.busy, Message := 'FullCycle#11 busy');
    AssertEquals_BOOL(Expected := FALSE, Actual := fbFullCycle.fault, Message := 'FullCycle#11 fault');
    AssertEquals_INT(Expected := 0, Actual := fbFullCycle.faultStep, Message := 'FullCycle#11 faultStep');
    AssertEquals_DINT(Expected := 1, Actual := fbFullCycle.cycleCount, Message := 'FullCycle#11 cycleCount');
    AssertEquals_STRING(Expected := 'IDLE', Actual := fbFullCycle.stepText, Message := 'FullCycle#11 stepText');

    GVL_S7Clock.xSimulation := FALSE;
END_IF
coUnit.TEST_FINISHED();

(* ---- PermissiveMissing.method.impl.st ---- *)
// AUTO-GENERATED — не редактировать: scenarios/FB_Sequencer.csv, сценарий PermissiveMissing
coUnit.TEST('PermissiveMissing');
IF NOT xPermissiveMissingDone THEN
    xPermissiveMissingDone := TRUE;
    GVL_S7Clock.xSimulation := TRUE;

    // #1, t = 0 мс — разрешения нет
    GVL_S7Clock.tSimNow := T#0MS;
    fbPermissiveMissing.start := FALSE;
    fbPermissiveMissing.stop := FALSE;
    fbPermissiveMissing.permissive := FALSE;
    fbPermissiveMissing.levelLow := FALSE;
    fbPermissiveMissing.levelHigh := FALSE;
    fbPermissiveMissing.reset := FALSE;
    fbPermissiveMissing.drainTimeout := T#60000MS;
    fbPermissiveMissing.airTime := T#30000MS;
    fbPermissiveMissing.washTime := T#40000MS;
    fbPermissiveMissing.refillTimeout := T#90000MS;
    fbPermissiveMissing();
    AssertEquals_INT(Expected := 0, Actual := fbPermissiveMissing.stepNo, Message := 'PermissiveMissing#1 stepNo');
    AssertEquals_BOOL(Expected := FALSE,
                      Actual := fbPermissiveMissing.drainValve,
                      Message := 'PermissiveMissing#1 drainValve');
    AssertEquals_BOOL(Expected := FALSE,
                      Actual := fbPermissiveMissing.airBlower,
                      Message := 'PermissiveMissing#1 airBlower');
    AssertEquals_BOOL(Expected := FALSE,
                      Actual := fbPermissiveMissing.washPump,
                      Message := 'PermissiveMissing#1 washPump');
    AssertEquals_BOOL(Expected := FALSE,
                      Actual := fbPermissiveMissing.inletValve,
                      Message := 'PermissiveMissing#1 inletValve');
    AssertEquals_BOOL(Expected := FALSE, Actual := fbPermissiveMissing.busy, Message := 'PermissiveMissing#1 busy');
    AssertEquals_BOOL(Expected := FALSE, Actual := fbPermissiveMissing.fault, Message := 'PermissiveMissing#1 fault');
    AssertEquals_INT(Expected := 0,
                     Actual := fbPermissiveMissing.faultStep,
                     Message := 'PermissiveMissing#1 faultStep');
    AssertEquals_DINT(Expected := 0,
                      Actual := fbPermissiveMissing.cycleCount,
                      Message := 'PermissiveMissing#1 cycleCount');
    AssertEquals_STRING(Expected := 'IDLE',
                        Actual := fbPermissiveMissing.stepText,
                        Message := 'PermissiveMissing#1 stepText');

    // #2, t = 1000 мс — фронт start без разрешения: ожидание
    GVL_S7Clock.tSimNow := T#1000MS;
    fbPermissiveMissing.start := TRUE;
    fbPermissiveMissing();
    AssertEquals_INT(Expected := 0, Actual := fbPermissiveMissing.stepNo, Message := 'PermissiveMissing#2 stepNo');
    AssertEquals_BOOL(Expected := FALSE,
                      Actual := fbPermissiveMissing.drainValve,
                      Message := 'PermissiveMissing#2 drainValve');
    AssertEquals_BOOL(Expected := FALSE,
                      Actual := fbPermissiveMissing.airBlower,
                      Message := 'PermissiveMissing#2 airBlower');
    AssertEquals_BOOL(Expected := FALSE,
                      Actual := fbPermissiveMissing.washPump,
                      Message := 'PermissiveMissing#2 washPump');
    AssertEquals_BOOL(Expected := FALSE,
                      Actual := fbPermissiveMissing.inletValve,
                      Message := 'PermissiveMissing#2 inletValve');
    AssertEquals_BOOL(Expected := FALSE, Actual := fbPermissiveMissing.busy, Message := 'PermissiveMissing#2 busy');
    AssertEquals_BOOL(Expected := FALSE, Actual := fbPermissiveMissing.fault, Message := 'PermissiveMissing#2 fault');
    AssertEquals_INT(Expected := 0,
                     Actual := fbPermissiveMissing.faultStep,
                     Message := 'PermissiveMissing#2 faultStep');
    AssertEquals_DINT(Expected := 0,
                      Actual := fbPermissiveMissing.cycleCount,
                      Message := 'PermissiveMissing#2 cycleCount');
    AssertEquals_STRING(Expected := 'IDLE',
                        Actual := fbPermissiveMissing.stepText,
                        Message := 'PermissiveMissing#2 stepText');

    // #3, t = 2000 мс — разрешение есть, start держится — фронта нет
    GVL_S7Clock.tSimNow := T#2000MS;
    fbPermissiveMissing.permissive := TRUE;
    fbPermissiveMissing();
    AssertEquals_INT(Expected := 0, Actual := fbPermissiveMissing.stepNo, Message := 'PermissiveMissing#3 stepNo');
    AssertEquals_BOOL(Expected := FALSE,
                      Actual := fbPermissiveMissing.drainValve,
                      Message := 'PermissiveMissing#3 drainValve');
    AssertEquals_BOOL(Expected := FALSE,
                      Actual := fbPermissiveMissing.airBlower,
                      Message := 'PermissiveMissing#3 airBlower');
    AssertEquals_BOOL(Expected := FALSE,
                      Actual := fbPermissiveMissing.washPump,
                      Message := 'PermissiveMissing#3 washPump');
    AssertEquals_BOOL(Expected := FALSE,
                      Actual := fbPermissiveMissing.inletValve,
                      Message := 'PermissiveMissing#3 inletValve');
    AssertEquals_BOOL(Expected := FALSE, Actual := fbPermissiveMissing.busy, Message := 'PermissiveMissing#3 busy');
    AssertEquals_BOOL(Expected := FALSE, Actual := fbPermissiveMissing.fault, Message := 'PermissiveMissing#3 fault');
    AssertEquals_INT(Expected := 0,
                     Actual := fbPermissiveMissing.faultStep,
                     Message := 'PermissiveMissing#3 faultStep');
    AssertEquals_DINT(Expected := 0,
                      Actual := fbPermissiveMissing.cycleCount,
                      Message := 'PermissiveMissing#3 cycleCount');
    AssertEquals_STRING(Expected := 'IDLE',
                        Actual := fbPermissiveMissing.stepText,
                        Message := 'PermissiveMissing#3 stepText');

    // #4, t = 3000 мс — start отпущен
    GVL_S7Clock.tSimNow := T#3000MS;
    fbPermissiveMissing.start := FALSE;
    fbPermissiveMissing();
    AssertEquals_INT(Expected := 0, Actual := fbPermissiveMissing.stepNo, Message := 'PermissiveMissing#4 stepNo');
    AssertEquals_BOOL(Expected := FALSE,
                      Actual := fbPermissiveMissing.drainValve,
                      Message := 'PermissiveMissing#4 drainValve');
    AssertEquals_BOOL(Expected := FALSE,
                      Actual := fbPermissiveMissing.airBlower,
                      Message := 'PermissiveMissing#4 airBlower');
    AssertEquals_BOOL(Expected := FALSE,
                      Actual := fbPermissiveMissing.washPump,
                      Message := 'PermissiveMissing#4 washPump');
    AssertEquals_BOOL(Expected := FALSE,
                      Actual := fbPermissiveMissing.inletValve,
                      Message := 'PermissiveMissing#4 inletValve');
    AssertEquals_BOOL(Expected := FALSE, Actual := fbPermissiveMissing.busy, Message := 'PermissiveMissing#4 busy');
    AssertEquals_BOOL(Expected := FALSE, Actual := fbPermissiveMissing.fault, Message := 'PermissiveMissing#4 fault');
    AssertEquals_INT(Expected := 0,
                     Actual := fbPermissiveMissing.faultStep,
                     Message := 'PermissiveMissing#4 faultStep');
    AssertEquals_DINT(Expected := 0,
                      Actual := fbPermissiveMissing.cycleCount,
                      Message := 'PermissiveMissing#4 cycleCount');
    AssertEquals_STRING(Expected := 'IDLE',
                        Actual := fbPermissiveMissing.stepText,
                        Message := 'PermissiveMissing#4 stepText');

    // #5, t = 4000 мс — новый фронт: опорожнение
    GVL_S7Clock.tSimNow := T#4000MS;
    fbPermissiveMissing.start := TRUE;
    fbPermissiveMissing();
    AssertEquals_INT(Expected := 10, Actual := fbPermissiveMissing.stepNo, Message := 'PermissiveMissing#5 stepNo');
    AssertEquals_BOOL(Expected := TRUE,
                      Actual := fbPermissiveMissing.drainValve,
                      Message := 'PermissiveMissing#5 drainValve');
    AssertEquals_BOOL(Expected := FALSE,
                      Actual := fbPermissiveMissing.airBlower,
                      Message := 'PermissiveMissing#5 airBlower');
    AssertEquals_BOOL(Expected := FALSE,
                      Actual := fbPermissiveMissing.washPump,
                      Message := 'PermissiveMissing#5 washPump');
    AssertEquals_BOOL(Expected := FALSE,
                      Actual := fbPermissiveMissing.inletValve,
                      Message := 'PermissiveMissing#5 inletValve');
    AssertEquals_BOOL(Expected := TRUE, Actual := fbPermissiveMissing.busy, Message := 'PermissiveMissing#5 busy');
    AssertEquals_BOOL(Expected := FALSE, Actual := fbPermissiveMissing.fault, Message := 'PermissiveMissing#5 fault');
    AssertEquals_INT(Expected := 0,
                     Actual := fbPermissiveMissing.faultStep,
                     Message := 'PermissiveMissing#5 faultStep');
    AssertEquals_DINT(Expected := 0,
                      Actual := fbPermissiveMissing.cycleCount,
                      Message := 'PermissiveMissing#5 cycleCount');
    AssertEquals_STRING(Expected := 'DRAIN',
                        Actual := fbPermissiveMissing.stepText,
                        Message := 'PermissiveMissing#5 stepText');

    GVL_S7Clock.xSimulation := FALSE;
END_IF
coUnit.TEST_FINISHED();

(* ---- RefillTimeoutBoundary.method.impl.st ---- *)
// AUTO-GENERATED — не редактировать: scenarios/FB_Sequencer.csv, сценарий RefillTimeoutBoundary
coUnit.TEST('RefillTimeoutBoundary');
IF NOT xRefillTimeoutBoundaryDone THEN
    xRefillTimeoutBoundaryDone := TRUE;
    GVL_S7Clock.xSimulation := TRUE;

    // #1, t = 0 мс — пуск: опорожнение; продувка и промывка по 5 с, заполнение до 10 с
    GVL_S7Clock.tSimNow := T#0MS;
    fbRefillTimeoutBoundary.start := TRUE;
    fbRefillTimeoutBoundary.stop := FALSE;
    fbRefillTimeoutBoundary.permissive := TRUE;
    fbRefillTimeoutBoundary.levelLow := FALSE;
    fbRefillTimeoutBoundary.levelHigh := FALSE;
    fbRefillTimeoutBoundary.reset := FALSE;
    fbRefillTimeoutBoundary.drainTimeout := T#60000MS;
    fbRefillTimeoutBoundary.airTime := T#5000MS;
    fbRefillTimeoutBoundary.washTime := T#5000MS;
    fbRefillTimeoutBoundary.refillTimeout := T#10000MS;
    fbRefillTimeoutBoundary();
    AssertEquals_INT(Expected := 10,
                     Actual := fbRefillTimeoutBoundary.stepNo,
                     Message := 'RefillTimeoutBoundary#1 stepNo');
    AssertEquals_BOOL(Expected := TRUE,
                      Actual := fbRefillTimeoutBoundary.drainValve,
                      Message := 'RefillTimeoutBoundary#1 drainValve');
    AssertEquals_BOOL(Expected := FALSE,
                      Actual := fbRefillTimeoutBoundary.airBlower,
                      Message := 'RefillTimeoutBoundary#1 airBlower');
    AssertEquals_BOOL(Expected := FALSE,
                      Actual := fbRefillTimeoutBoundary.washPump,
                      Message := 'RefillTimeoutBoundary#1 washPump');
    AssertEquals_BOOL(Expected := FALSE,
                      Actual := fbRefillTimeoutBoundary.inletValve,
                      Message := 'RefillTimeoutBoundary#1 inletValve');
    AssertEquals_BOOL(Expected := TRUE,
                      Actual := fbRefillTimeoutBoundary.busy,
                      Message := 'RefillTimeoutBoundary#1 busy');
    AssertEquals_BOOL(Expected := FALSE,
                      Actual := fbRefillTimeoutBoundary.fault,
                      Message := 'RefillTimeoutBoundary#1 fault');
    AssertEquals_INT(Expected := 0,
                     Actual := fbRefillTimeoutBoundary.faultStep,
                     Message := 'RefillTimeoutBoundary#1 faultStep');
    AssertEquals_DINT(Expected := 0,
                      Actual := fbRefillTimeoutBoundary.cycleCount,
                      Message := 'RefillTimeoutBoundary#1 cycleCount');
    AssertEquals_STRING(Expected := 'DRAIN',
                        Actual := fbRefillTimeoutBoundary.stepText,
                        Message := 'RefillTimeoutBoundary#1 stepText');

    // #2, t = 1000 мс — продувка с 1.0 с
    GVL_S7Clock.tSimNow := T#1000MS;
    fbRefillTimeoutBoundary.start := FALSE;
    fbRefillTimeoutBoundary.levelLow := TRUE;
    fbRefillTimeoutBoundary();
    AssertEquals_INT(Expected := 20,
                     Actual := fbRefillTimeoutBoundary.stepNo,
                     Message := 'RefillTimeoutBoundary#2 stepNo');
    AssertEquals_BOOL(Expected := FALSE,
                      Actual := fbRefillTimeoutBoundary.drainValve,
                      Message := 'RefillTimeoutBoundary#2 drainValve');
    AssertEquals_BOOL(Expected := TRUE,
                      Actual := fbRefillTimeoutBoundary.airBlower,
                      Message := 'RefillTimeoutBoundary#2 airBlower');
    AssertEquals_BOOL(Expected := FALSE,
                      Actual := fbRefillTimeoutBoundary.washPump,
                      Message := 'RefillTimeoutBoundary#2 washPump');
    AssertEquals_BOOL(Expected := FALSE,
                      Actual := fbRefillTimeoutBoundary.inletValve,
                      Message := 'RefillTimeoutBoundary#2 inletValve');
    AssertEquals_BOOL(Expected := TRUE,
                      Actual := fbRefillTimeoutBoundary.busy,
                      Message := 'RefillTimeoutBoundary#2 busy');
    AssertEquals_BOOL(Expected := FALSE,
                      Actual := fbRefillTimeoutBoundary.fault,
                      Message := 'RefillTimeoutBoundary#2 fault');
    AssertEquals_INT(Expected := 0,
                     Actual := fbRefillTimeoutBoundary.faultStep,
                     Message := 'RefillTimeoutBoundary#2 faultStep');
    AssertEquals_DINT(Expected := 0,
                      Actual := fbRefillTimeoutBoundary.cycleCount,
                      Message := 'RefillTimeoutBoundary#2 cycleCount');
    AssertEquals_STRING(Expected := 'AIR SCOUR',
                        Actual := fbRefillTimeoutBoundary.stepText,
                        Message := 'RefillTimeoutBoundary#2 stepText');

    // #3, t = 6400 мс — 5.4 с: промывка с 6.4 с
    GVL_S7Clock.tSimNow := T#6400MS;
    fbRefillTimeoutBoundary.levelLow := FALSE;
    fbRefillTimeoutBoundary();
    AssertEquals_INT(Expected := 30,
                     Actual := fbRefillTimeoutBoundary.stepNo,
                     Message := 'RefillTimeoutBoundary#3 stepNo');
    AssertEquals_BOOL(Expected := TRUE,
                      Actual := fbRefillTimeoutBoundary.drainValve,
                      Message := 'RefillTimeoutBoundary#3 drainValve');
    AssertEquals_BOOL(Expected := FALSE,
                      Actual := fbRefillTimeoutBoundary.airBlower,
                      Message := 'RefillTimeoutBoundary#3 airBlower');
    AssertEquals_BOOL(Expected := TRUE,
                      Actual := fbRefillTimeoutBoundary.washPump,
                      Message := 'RefillTimeoutBoundary#3 washPump');
    AssertEquals_BOOL(Expected := FALSE,
                      Actual := fbRefillTimeoutBoundary.inletValve,
                      Message := 'RefillTimeoutBoundary#3 inletValve');
    AssertEquals_BOOL(Expected := TRUE,
                      Actual := fbRefillTimeoutBoundary.busy,
                      Message := 'RefillTimeoutBoundary#3 busy');
    AssertEquals_BOOL(Expected := FALSE,
                      Actual := fbRefillTimeoutBoundary.fault,
                      Message := 'RefillTimeoutBoundary#3 fault');
    AssertEquals_INT(Expected := 0,
                     Actual := fbRefillTimeoutBoundary.faultStep,
                     Message := 'RefillTimeoutBoundary#3 faultStep');
    AssertEquals_DINT(Expected := 0,
                      Actual := fbRefillTimeoutBoundary.cycleCount,
                      Message := 'RefillTimeoutBoundary#3 cycleCount');
    AssertEquals_STRING(Expected := 'BACKWASH',
                        Actual := fbRefillTimeoutBoundary.stepText,
                        Message := 'RefillTimeoutBoundary#3 stepText');

    // #4, t = 11800 мс — 5.4 с: заполнение с 11.8 с
    GVL_S7Clock.tSimNow := T#11800MS;
    fbRefillTimeoutBoundary();
    AssertEquals_INT(Expected := 40,
                     Actual := fbRefillTimeoutBoundary.stepNo,
                     Message := 'RefillTimeoutBoundary#4 stepNo');
    AssertEquals_BOOL(Expected := FALSE,
                      Actual := fbRefillTimeoutBoundary.drainValve,
                      Message := 'RefillTimeoutBoundary#4 drainValve');
    AssertEquals_BOOL(Expected := FALSE,
                      Actual := fbRefillTimeoutBoundary.airBlower,
                      Message := 'RefillTimeoutBoundary#4 airBlower');
    AssertEquals_BOOL(Expected := FALSE,
                      Actual := fbRefillTimeoutBoundary.washPump,
                      Message := 'RefillTimeoutBoundary#4 washPump');
    AssertEquals_BOOL(Expected := TRUE,
                      Actual := fbRefillTimeoutBoundary.inletValve,
                      Message := 'RefillTimeoutBoundary#4 inletValve');
    AssertEquals_BOOL(Expected := TRUE,
                      Actual := fbRefillTimeoutBoundary.busy,
                      Message := 'RefillTimeoutBoundary#4 busy');
    AssertEquals_BOOL(Expected := FALSE,
                      Actual := fbRefillTimeoutBoundary.fault,
                      Message := 'RefillTimeoutBoundary#4 fault');
    AssertEquals_INT(Expected := 0,
                     Actual := fbRefillTimeoutBoundary.faultStep,
                     Message := 'RefillTimeoutBoundary#4 faultStep');
    AssertEquals_DINT(Expected := 0,
                      Actual := fbRefillTimeoutBoundary.cycleCount,
                      Message := 'RefillTimeoutBoundary#4 cycleCount');
    AssertEquals_STRING(Expected := 'REFILL',
                        Actual := fbRefillTimeoutBoundary.stepText,
                        Message := 'RefillTimeoutBoundary#4 stepText');

    // #5, t = 21600 мс — 9.8 с < 10 с: заполнение
    GVL_S7Clock.tSimNow := T#21600MS;
    fbRefillTimeoutBoundary();
    AssertEquals_INT(Expected := 40,
                     Actual := fbRefillTimeoutBoundary.stepNo,
                     Message := 'RefillTimeoutBoundary#5 stepNo');
    AssertEquals_BOOL(Expected := FALSE,
                      Actual := fbRefillTimeoutBoundary.drainValve,
                      Message := 'RefillTimeoutBoundary#5 drainValve');
    AssertEquals_BOOL(Expected := FALSE,
                      Actual := fbRefillTimeoutBoundary.airBlower,
                      Message := 'RefillTimeoutBoundary#5 airBlower');
    AssertEquals_BOOL(Expected := FALSE,
                      Actual := fbRefillTimeoutBoundary.washPump,
                      Message := 'RefillTimeoutBoundary#5 washPump');
    AssertEquals_BOOL(Expected := TRUE,
                      Actual := fbRefillTimeoutBoundary.inletValve,
                      Message := 'RefillTimeoutBoundary#5 inletValve');
    AssertEquals_BOOL(Expected := TRUE,
                      Actual := fbRefillTimeoutBoundary.busy,
                      Message := 'RefillTimeoutBoundary#5 busy');
    AssertEquals_BOOL(Expected := FALSE,
                      Actual := fbRefillTimeoutBoundary.fault,
                      Message := 'RefillTimeoutBoundary#5 fault');
    AssertEquals_INT(Expected := 0,
                     Actual := fbRefillTimeoutBoundary.faultStep,
                     Message := 'RefillTimeoutBoundary#5 faultStep');
    AssertEquals_DINT(Expected := 0,
                      Actual := fbRefillTimeoutBoundary.cycleCount,
                      Message := 'RefillTimeoutBoundary#5 cycleCount');
    AssertEquals_STRING(Expected := 'REFILL',
                        Actual := fbRefillTimeoutBoundary.stepText,
                        Message := 'RefillTimeoutBoundary#5 stepText');

    // #6, t = 21800 мс, на пороге таймера — 10.0 с = refillTimeout: авария на шаге 40
    GVL_S7Clock.tSimNow := T#21800MS;
    fbRefillTimeoutBoundary();
    AssertEquals_INT(Expected := 90,
                     Actual := fbRefillTimeoutBoundary.stepNo,
                     Message := 'RefillTimeoutBoundary#6 stepNo');
    AssertEquals_BOOL(Expected := FALSE,
                      Actual := fbRefillTimeoutBoundary.drainValve,
                      Message := 'RefillTimeoutBoundary#6 drainValve');
    AssertEquals_BOOL(Expected := FALSE,
                      Actual := fbRefillTimeoutBoundary.airBlower,
                      Message := 'RefillTimeoutBoundary#6 airBlower');
    AssertEquals_BOOL(Expected := FALSE,
                      Actual := fbRefillTimeoutBoundary.washPump,
                      Message := 'RefillTimeoutBoundary#6 washPump');
    AssertEquals_BOOL(Expected := FALSE,
                      Actual := fbRefillTimeoutBoundary.inletValve,
                      Message := 'RefillTimeoutBoundary#6 inletValve');
    AssertEquals_BOOL(Expected := FALSE,
                      Actual := fbRefillTimeoutBoundary.busy,
                      Message := 'RefillTimeoutBoundary#6 busy');
    AssertEquals_BOOL(Expected := TRUE,
                      Actual := fbRefillTimeoutBoundary.fault,
                      Message := 'RefillTimeoutBoundary#6 fault');
    AssertEquals_INT(Expected := 40,
                     Actual := fbRefillTimeoutBoundary.faultStep,
                     Message := 'RefillTimeoutBoundary#6 faultStep');
    AssertEquals_DINT(Expected := 0,
                      Actual := fbRefillTimeoutBoundary.cycleCount,
                      Message := 'RefillTimeoutBoundary#6 cycleCount');
    AssertEquals_STRING(Expected := 'FAULT',
                        Actual := fbRefillTimeoutBoundary.stepText,
                        Message := 'RefillTimeoutBoundary#6 stepText');

    // #7, t = 22000 мс — авария
    GVL_S7Clock.tSimNow := T#22000MS;
    fbRefillTimeoutBoundary();
    AssertEquals_INT(Expected := 90,
                     Actual := fbRefillTimeoutBoundary.stepNo,
                     Message := 'RefillTimeoutBoundary#7 stepNo');
    AssertEquals_BOOL(Expected := FALSE,
                      Actual := fbRefillTimeoutBoundary.drainValve,
                      Message := 'RefillTimeoutBoundary#7 drainValve');
    AssertEquals_BOOL(Expected := FALSE,
                      Actual := fbRefillTimeoutBoundary.airBlower,
                      Message := 'RefillTimeoutBoundary#7 airBlower');
    AssertEquals_BOOL(Expected := FALSE,
                      Actual := fbRefillTimeoutBoundary.washPump,
                      Message := 'RefillTimeoutBoundary#7 washPump');
    AssertEquals_BOOL(Expected := FALSE,
                      Actual := fbRefillTimeoutBoundary.inletValve,
                      Message := 'RefillTimeoutBoundary#7 inletValve');
    AssertEquals_BOOL(Expected := FALSE,
                      Actual := fbRefillTimeoutBoundary.busy,
                      Message := 'RefillTimeoutBoundary#7 busy');
    AssertEquals_BOOL(Expected := TRUE,
                      Actual := fbRefillTimeoutBoundary.fault,
                      Message := 'RefillTimeoutBoundary#7 fault');
    AssertEquals_INT(Expected := 40,
                     Actual := fbRefillTimeoutBoundary.faultStep,
                     Message := 'RefillTimeoutBoundary#7 faultStep');
    AssertEquals_DINT(Expected := 0,
                      Actual := fbRefillTimeoutBoundary.cycleCount,
                      Message := 'RefillTimeoutBoundary#7 cycleCount');
    AssertEquals_STRING(Expected := 'FAULT',
                        Actual := fbRefillTimeoutBoundary.stepText,
                        Message := 'RefillTimeoutBoundary#7 stepText');

    // #8, t = 23000 мс — сброс
    GVL_S7Clock.tSimNow := T#23000MS;
    fbRefillTimeoutBoundary.reset := TRUE;
    fbRefillTimeoutBoundary();
    AssertEquals_INT(Expected := 0,
                     Actual := fbRefillTimeoutBoundary.stepNo,
                     Message := 'RefillTimeoutBoundary#8 stepNo');
    AssertEquals_BOOL(Expected := FALSE,
                      Actual := fbRefillTimeoutBoundary.drainValve,
                      Message := 'RefillTimeoutBoundary#8 drainValve');
    AssertEquals_BOOL(Expected := FALSE,
                      Actual := fbRefillTimeoutBoundary.airBlower,
                      Message := 'RefillTimeoutBoundary#8 airBlower');
    AssertEquals_BOOL(Expected := FALSE,
                      Actual := fbRefillTimeoutBoundary.washPump,
                      Message := 'RefillTimeoutBoundary#8 washPump');
    AssertEquals_BOOL(Expected := FALSE,
                      Actual := fbRefillTimeoutBoundary.inletValve,
                      Message := 'RefillTimeoutBoundary#8 inletValve');
    AssertEquals_BOOL(Expected := FALSE,
                      Actual := fbRefillTimeoutBoundary.busy,
                      Message := 'RefillTimeoutBoundary#8 busy');
    AssertEquals_BOOL(Expected := FALSE,
                      Actual := fbRefillTimeoutBoundary.fault,
                      Message := 'RefillTimeoutBoundary#8 fault');
    AssertEquals_INT(Expected := 0,
                     Actual := fbRefillTimeoutBoundary.faultStep,
                     Message := 'RefillTimeoutBoundary#8 faultStep');
    AssertEquals_DINT(Expected := 0,
                      Actual := fbRefillTimeoutBoundary.cycleCount,
                      Message := 'RefillTimeoutBoundary#8 cycleCount');
    AssertEquals_STRING(Expected := 'IDLE',
                        Actual := fbRefillTimeoutBoundary.stepText,
                        Message := 'RefillTimeoutBoundary#8 stepText');

    GVL_S7Clock.xSimulation := FALSE;
END_IF
coUnit.TEST_FINISHED();
